(* IEC 61131-3 sources: codesys-to-s7/tests/corpus/C2S7-TYPE-STRLEN/pos, 1 file *)

(* ---- input.st ---- *)
FUNCTION_BLOCK FB_Case
VAR
    s : STRING(300);
END_VAR
s := 'a';
END_FUNCTION_BLOCK
